(* CODESYS project keyence_iv.library
   Company: KOSTAL GmbH & Co.KG
   Version: 2.0.0.0
   DefaultNamespace: KOSTAL.AF2024.Drivers.Camera.Keyence_IV
   Title: KOSTAL.AF2024.Drivers.Camera.Keyence_IV
   Placeholder: KOSTAL.AF2024.Drivers.Camera.Keyence_IV
   Author: Frank Dümpelmann, Martin Hundt
   DocFormat: reStructuredText

Project tree, tasks and I/O mapping:
  libraries: KOSTAL.AF2024.Core.functionResponse, 1.0.0.0 (KOSTAL GmbH & Co.KG); KOSTAL.AF2024.Core.ListOf, 1.0.0.0 (KOSTAL GmbH & Co.KG); KOSTAL.AF2024.Core.Process, 1.0.0.0 (KOSTAL GmbH & Co.KG); KOSTAL.AF2024.Core.Settings, 1.0.0.0 (KOSTAL GmbH & Co.KG); KOSTAL.AF2024.Core.StringTools, 1.0.0.0 (KOSTAL GmbH & Co.KG); KOSTAL.AF2024.Core.System, 1.0.0.0 (KOSTAL GmbH & Co.KG); KOSTAL.AF2024.Drivers.Camera.I_Camera, 2.0.0.0 (KOSTAL GmbH & Co.KG); Tc2_Standard, 3.3.3.0 (Beckhoff Automation GmbH); Tc2_System, 3.6.2.0 (Beckhoff Automation GmbH); Tc2_TcpIp, 3.3.10.0 (Beckhoff Automation GmbH)
  DIO/
    DUT/
      data type _E_PROCESS
      data type _ST_fromDevice
      data type _ST_fromDevice_HG_
      data type _ST_toDevice
    function block FB_Camera_DIO_IV [ST]: Ex_SetProgramNumber, Ex_Trigger, Ex_Trigger_ProgramNumber, ProgramNumber, ResultPass, State, _setFinish, _toDevice_Clear, _faultHandler, _fbMain, _idle, _sequence, _setProgram, Fault, FaultReset, FBmain
    function block FB_Camera_DIO_IV_HG [ST]: CustomOut_5, CustomOut_6, CustomOut_7, CustomOut_8
  Project Information/
    function F_GetCompany [ST]
    function F_GetTitle [ST]
    function F_GetVersion [ST]
  TcpIp/
    DUT/
      _Internal/
        data type _E_Command_TcpIp
        data type _E_THIS_TcpIp
        function block _T_Command [ST]: Error, GetProgram, OK, ReadOperationMode, ReadVersion, SetProgram, StateResult, TriggerAndState
      Response RT/
        interface I_T_Response_RT_TcpIp: CopyTo, OverallPass, ResultCount, Tools
        interface I_T_Response_RT_TcpIp_CopyFrom: CopyFrom
        interface I_T_Response_RT_TcpIp_Owner: Clear, CopyFrom, OverallPass, ResultCount, Tools_Owner
        function block T_Response_RT_TcpIp [ST]: Clear, CopyFrom, CopyTo, OverallPass, ResultCount, Tools, Tools_Owner
      Tool/
        ListOf/
          function block FB_ListOf_T_Tool [ST]: _get_I, _get_I_Owner, _removePayLoad, _verifyMember, Add_DUT, Clear, CopyFrom, CopyTo, Delete_DUT, Get_I, Get_I_Owner, NumberOfMember
          interface I_ListOf_T_Tool: CopyTo, Get_I, NumberOfMember
          interface I_ListOf_T_Tool_CopyFrom: CopyFrom
          interface I_ListOf_T_Tool_Owner: Add_DUT, Clear, CopyFrom, CopyTo, Delete_DUT, Get_I, Get_I_Owner, NumberOfMember
        interface I_T_Tool: CopyTo, MatchingRate, Number, Pass
        interface I_T_Tool_CopyFrom: CopyFrom
        interface I_T_Tool_Owner: Clear, CopyFrom, MatchingRate, Number, Pass
        function block T_Tool [ST]: Clear, CopyFrom, CopyTo, MatchingRate, Number, Pass
      Version/
        interface I_T_SensorVersion_TcpIp: CopyTo, HeadModel, Version
        interface I_T_SensorVersion_TcpIp_CopyFrom: CopyFrom
        interface I_T_SensorVersion_TcpIp_Owner: Clear, CopyFrom, HeadModel, Version
        function block T_SensorVersion_TcpIp [ST]: Clear, CopyFrom, CopyTo, HeadModel, Version
      data type E_OpMode_TcpIp
    function block FB_Camera_TcpIp_IV [ST]: FB_init, _getCommand, _mergePlCommand, _Parse_Error, _Parse_ErrorMessage, _Parse_GetProgram, _Parse_OpMode, _Parse_SetProgram, _Parse_Trigger, _Parse_Version, _a0_stepFail, _a0_stepInit, _a1_Finish, _a1_Idle, _a2_Connect, _a2_Parse, _a2_Receive, _a2_Send, _a3_PrgIsEqual, _devices, _splitString, _timeOutOccured, _FBmain, Clear, Ex_GetProgramNumber, Ex_ReadOperationMode, Ex_ReadVersion, Ex_SetProgramNumber, Ex_Trigger, Ex_Trigger_ProgramNumber, GetElement, NativeStringGet, IP, Port, Content, ExecutedSocketState, NumberOfEntries, OperationMode, Result, ResultPass, serverAmsNetId, State, Version, FBmain
    interface I_Camera_TcpIp_IV: GetElement, NativeStringGet, Content, ExecutedSocketState, IP, NumberOfEntries, OperationMode, Port, Result, serverAmsNetId
  Version/
    global variables Global_Version
*)

// DIO/DUT/_E_PROCESS
{attribute 'qualified_only'}
{attribute 'strict'}
TYPE _E_PROCESS :
(
	idle		:= 0,
	Start		:= 1, 
	SetProgram	:= 2
);
END_TYPE

// DIO/DUT/_ST_fromDevice
TYPE _ST_fromDevice :
STRUCT
	TotalStatusOK	:BOOL;
	Busy			:BOOL;
	Error			:BOOL;
	Run				:BOOL;
END_STRUCT
END_TYPE

// DIO/DUT/_ST_fromDevice_HG_
TYPE _ST_fromDevice_HG_ :
STRUCT
	CustomOut_5		: BOOL;
	CustomOut_6		: BOOL;
	CustomOut_7		: BOOL;
	CustomOut_8		: BOOL;
END_STRUCT
END_TYPE

// DIO/DUT/_ST_toDevice
TYPE _ST_toDevice:
	STRUCT
		ExternalTrigger		:BOOL;
		ProgramSelectBit0	:BOOL;
		ProgramSelectBit1	:BOOL;
		ProgramSelectBit2	:BOOL;
		ProgramSelectBit3	:BOOL;
		ErrorClear			:BOOL;
	END_STRUCT
END_TYPE

// TcpIp/DUT/_Internal/_E_Command_TcpIp
{attribute 'qualified_only'}
{attribute 'strict'}
TYPE INTERNAL _E_Command_TcpIp :
(
	Trigger := 0,
	SetProgram,
	GetProgram,
	ReadVersion,
	ReadOperationMode
);
END_TYPE

// TcpIp/DUT/_Internal/_E_THIS_TcpIp
{attribute 'qualified_only'}
{attribute 'strict'}
TYPE INTERNAL _E_THIS_TcpIp :
(
	Idle := 0,
	Trigger,
	TriggerPrgNo,
	SetProgram,
	GetProgram,
	ReadVersion,
	ReadOperationMode
);
END_TYPE

// TcpIp/DUT/E_OpMode_TcpIp
{attribute 'qualified_only'}
{attribute 'strict'}
TYPE E_OpMode_TcpIp :
(
	Unknown := 0,
	Setup,
	Run
);
END_TYPE

// Version/Global_Version
{attribute 'TcGenerated'}
{attribute 'no-analysis'}
{attribute 'linkalways'}
// This function has been automatically generated from the project information.
VAR_GLOBAL CONSTANT
	{attribute 'const_non_replaced'}
	stLibVersion_KOSTAL_AF2024_Drivers_Camera_Keyence_IV : ST_LibVersion := (iMajor := 2, iMinor := 0, iBuild := 0, iRevision := 0, nFlags := 0, sVersion := '2.0.0.0');
END_VAR

// DIO/FB_Camera_DIO_IV
(*

:Author: Martin Hundt <m.hundt@kostal.com>
:Date: 2022-03-11

Function
========
| Device driver for Keyence IV-Series vision sensors with discrete IOs
| Selection of 15 sensor programs (program No. 0 is reserved)

Methods and Properties
======================
| Ex_start: Start the last selected camera program
| Ex_start_ProgramNumber: Start the camera program number in the method's parameter (int)

| State.ready: Camera is ready
| State.busy: Camera is analysing an image
| State.finish: Image analysis was finished
| State.pass: Image was processed -> Check result
| State.fail: Image image processing failed

| Fault: Camera in error state


Sensor Configuration
=====================
| The following IOs must be configured at the sensor and linked to the hardware IOs according to their names:
| Sensor Outputs: TotalStatusOK, Busy, Error, Run				
| Sensor Inputs: ExternalTrigger, ProgramSelectBit0, ProgramSelectBit1, ProgramSelectBit2, ErrorClear			

*)

FUNCTION_BLOCK FB_Camera_DIO_IV IMPLEMENTS KOSTAL_AF2024_Drivers_Camera_I_Camera.I_CameraWithFeedback
VAR
	_fromSensor AT %I*	: _ST_fromDevice;
	_toSensor 	AT %Q*	: _ST_toDevice;
	
	_THIS_CALLED		: _E_PROCESS;
	_THIS_IN_PROCESS	: _E_PROCESS;
	_step				: KOSTAL_AF2024_Core_Process.FB_processStep;
	_state				: KOSTAL_AF2024_Core_Process.T_plcState;
	
	_programNoOld		: USINT;
	_init				: BOOL;		(*BOOL - initialization required*)
	_triggerBusy		: F_TRIG;	(*F_TRIG*)
	_responseTime		: TON;	(*TON*)
	_resetClock			: TP;		(*TP*)
	
	_faultReset			: BOOL;
	
	_resultPass			: BOOL;
	_resultFail			: BOOL;
	
	_programNo			: USINT;
	_fault				: BOOL;
	                    
END_VAR

METHOD Ex_SetProgramNumber : BOOL;
VAR_INPUT
	ProgramNumber	: UINT;
END_VAR
IF _THIS_CALLED <> _E_PROCESS.idle THEN //Another process is running: don't start this process!
	Ex_SetProgramNumber:= FALSE;	
	RETURN; 
END_IF

_programNo := UINT_TO_USINT(ProgramNumber);
_THIS_CALLED := _E_PROCESS.SetProgram;

_FBmain();	//Call sequence via _FBmain

Ex_SetProgramNumber := _THIS_CALLED = _THIS_IN_PROCESS;	//Return true when process was started
END_METHOD

METHOD Ex_Trigger : BOOL;
IF _THIS_CALLED <> _E_PROCESS.idle THEN //Another process is running: don't start this process!
	Ex_Trigger:= FALSE;	
	RETURN; 
END_IF


_THIS_CALLED := _E_PROCESS.Start;

_FBmain();	//Call sequence via _FBmain

Ex_Trigger := _THIS_CALLED = _THIS_IN_PROCESS;	//Return true when process was started
END_METHOD

METHOD Ex_Trigger_ProgramNumber : BOOL;
VAR_INPUT
	ProgramNumber	: UINT;
END_VAR
IF _THIS_CALLED <> _E_PROCESS.idle THEN //Another process is running: don't start this process!
	Ex_Trigger_ProgramNumber:= FALSE;	
	RETURN; 
END_IF

_programNo := UINT_TO_USINT(ProgramNumber);
_THIS_CALLED := _E_PROCESS.Start;

_FBmain();	//Call sequence via _FBmain

Ex_Trigger_ProgramNumber := _THIS_CALLED = _THIS_IN_PROCESS;	//Return true when process was started
END_METHOD

PROPERTY PUBLIC ProgramNumber : UINT
GET
ProgramNumber := _programNo;
END_GET
END_PROPERTY

PROPERTY PUBLIC ResultPass : BOOL
GET
ResultPass := _resultPass;
END_GET
END_PROPERTY

PROPERTY State : KOSTAL_AF2024_Core_Process.I_T_plcState
GET

State := _state;
END_GET
END_PROPERTY

METHOD PROTECTED _setFinish
VAR_INPUT
END_VAR
END_METHOD

METHOD PROTECTED _toDevice_Clear
VAR_INPUT
END_VAR
_toSensor.ErrorClear := FALSE;
_toSensor.ExternalTrigger := FALSE;
_toSensor.ProgramSelectBit0 := FALSE;
_toSensor.ProgramSelectBit1 := FALSE;
_toSensor.ProgramSelectBit2 := FALSE;
_toSensor.ProgramSelectBit3 := FALSE;
END_METHOD

METHOD PROTECTED _faultHandler : BOOL
VAR_INPUT
END_VAR
_fault:= _fromSensor.Error;

IF _fromSensor.Error THEN
	_state.clear();
	_state.Fail:= TRUE;
	_state.Description:= "Device send >ERROR<";	
	
	_toDevice_Clear();

	_resetClock(IN:= _faultReset, PT:= T#250MS);
	_toSensor.ErrorClear:= _resetClock.Q;	
ELSE
	_faultHandler := TRUE;
END_IF

_faultReset := false;
END_METHOD

METHOD Protected _fbMain
VAR_INPUT
END_VAR
IF NOT _init THEN
	_step.init();
	_programNoOld:= 0;
	_resetClock(IN:= FALSE);
	_init:= TRUE;
	_toDevice_Clear();
END_IF

IF NOT _faultHandler() THEN RETURN; END_IF


IF _THIS_CALLED <> _THIS_IN_PROCESS THEN
	_step.init();
END_IF

_THIS_IN_PROCESS:= _THIS_CALLED;

CASE _THIS_CALLED OF
	_E_PROCESS.SetProgram:
		_setProgram();
	_E_PROCESS.Start:
		_sequence();
ELSE
	_idle();
END_CASE
END_METHOD

METHOD PROTECTED _idle
VAR_INPUT
END_VAR
_step.init();

_toSensor.ErrorClear:= FALSE;
_toSensor.ExternalTrigger := FALSE;
_resultPass := FALSE;
_resultFail := FALSE;
_state.clear();
_state.Ready := TRUE;
END_METHOD

METHOD PROTECTED _sequence
VAR_INPUT
END_VAR
_step.Header();

CASE _step.actual OF		
	0: //Check Program No.
		_state.clear();
		_state.Busy := TRUE;
		IF (_programNo = 0) OR (_programNo > 15) THEN
			_state.clear();
			_state.finish:= TRUE;
			_state.Fail:= TRUE;
			_state.Description:= "ProgramNo out of range (1<Pno>15)";
		ELSE
			_step.INC();
		END_IF

	1: (*Change Program *)
		IF _step.Toggle THEN
			_responseTime(IN:= FALSE);
			_triggerBusy(CLK:= FALSE);
		END_IF

		_toSensor.ProgramSelectBit0 := _programNo.0;
		_toSensor.ProgramSelectBit1 := _programNo.1;
		_toSensor.ProgramSelectBit2 := _programNo.2;
		_toSensor.ProgramSelectBit3 := _programNo.3;

		_state.clear();
		_state.Busy := TRUE;
		_state.Description:= "send program Number";

		_responseTime(IN:= TRUE, PT:= T#1s);
		_triggerBusy(CLK:=_fromSensor.Busy);	(*Wait until program is changed*)

		IF _programNo <> _programNoOld THEN

			IF _triggerBusy.Q OR _responseTime.Q THEN
				_programNoOld := _programNo;
			END_IF

		ELSE
			_step.INC();
		END_IF

	2:	(*trigger*)
		_toSensor.ExternalTrigger := TRUE;

		_state.clear();
		_state.Busy := TRUE;
		_state.Description:= "wait sensor busy";

		IF NOT _fromSensor.Run THEN
			_state.clear();
			_state.finish := TRUE;
			_state.fail := TRUE;
			_state.Description:= "Device not in >RUN<";
		ELSIF _fromSensor.Busy THEN
			_step.INC();
		END_IF

	3:	(*Read result*)
		_toSensor.ExternalTrigger := TRUE;

		_state.clear();
		_state.Busy := TRUE;
		_state.Description:=  "wait sensor finish";

		IF NOT _fromSensor.Busy THEN
			_step.INC();
		END_IF

	4:	(*finish*)
		_toSensor.ExternalTrigger := TRUE;
		_state.clear();
		_state.Finish := TRUE;
		_state.pass := TRUE;
		
		_resultPass:= _fromSensor.TotalStatusOK;
		_resultFail:= NOT _fromSensor.TotalStatusOK;

		
		IF _resultPass THEN
			_state.Description:= "get PASS";
		ELSE
			_state.Description:= "get FAIL";
		END_IF
		

END_CASE
END_METHOD

METHOD PROTECTED _setProgram
VAR_INPUT
END_VAR
_state.clear();
IF (_programNo = 0) OR (_programNo > 15) THEN
	_state.finish:= TRUE;
	_state.Fail:= TRUE;
	_state.Description:= "ProgramNo out of range (1<Pno>15)";
ELSE
	_state.finish:= TRUE;
	_state.pass:= TRUE;
END_IF
END_METHOD

PROPERTY Fault : BOOL
GET
Fault := _fault;
END_GET
END_PROPERTY

METHOD PUBLIC FaultReset
VAR_INPUT
END_VAR
_faultReset := True;
END_METHOD

METHOD PUBLIC FBmain
VAR_INPUT
END_VAR
IF _THIS_CALLED = _E_PROCESS.idle THEN
	
	_FBmain();
	
END_IF

_THIS_CALLED:= _E_PROCESS.idle;
END_METHOD

END_FUNCTION_BLOCK

// DIO/FB_Camera_DIO_IV_HG
//Extension of FB_Camera_IV with four custom outputs (only available for IV-HG device)
FUNCTION_BLOCK FB_Camera_DIO_IV_HG EXTENDS FB_Camera_DIO_IV
VAR
	_fromdeviceCustom	AT %I*	: _ST_fromDevice_HG_;
END_VAR

PROPERTY PUBLIC CustomOut_5 : Bool
GET
CustomOut_5 := _fromdeviceCustom.CustomOut_5;
END_GET
END_PROPERTY

PROPERTY PUBLIC CustomOut_6 : Bool
GET
CustomOut_6 := _fromdeviceCustom.CustomOut_6;
END_GET
END_PROPERTY

PROPERTY PUBLIC CustomOut_7 : Bool
GET
CustomOut_7 := _fromdeviceCustom.CustomOut_7;
END_GET
END_PROPERTY

PROPERTY PUBLIC CustomOut_8 : Bool
GET
CustomOut_8 := _fromdeviceCustom.CustomOut_8;
END_GET
END_PROPERTY

END_FUNCTION_BLOCK

// Project Information/F_GetCompany
// This function has been automatically generated from the project information.
{attribute 'signature_flag' := '1073741824'}
{attribute 'TcGenerated'}
{attribute 'no-analysis'}
FUNCTION F_GetCompany : WSTRING
VAR_INPUT
	
END_VAR

F_GetCompany := "KOSTAL GmbH & Co.KG";

END_FUNCTION

// Project Information/F_GetTitle
// This function has been automatically generated from the project information.
{attribute 'signature_flag' := '1073741824'}
{attribute 'TcGenerated'}
{attribute 'no-analysis'}
FUNCTION F_GetTitle : WSTRING
VAR_INPUT
	
END_VAR

F_GetTitle := "KOSTAL.AF2024.Drivers.Camera.Keyence_IV";

END_FUNCTION

// Project Information/F_GetVersion
// This function has been automatically generated from the project information.
{attribute 'signature_flag' := '1073741824'}
{attribute 'TcGenerated'}
{attribute 'no-analysis'}
FUNCTION F_GetVersion : ST_LibVersion
VAR_INPUT
	
END_VAR

F_GetVersion.iMajor := 2;
F_GetVersion.iMinor := 0;
F_GetVersion.iBuild := 0;
F_GetVersion.iRevision := 0;
F_GetVersion.sVersion := '2.0.0.0';
F_GetVersion.nFlags := 0;

END_FUNCTION

// TcpIp/DUT/_Internal/_T_Command
FUNCTION_BLOCK INTERNAL _T_Command

PROPERTY PUBLIC Error : STRING
GET

Error	:= 'ER';
END_GET
END_PROPERTY

PROPERTY PUBLIC GetProgram : STRING
GET

GetProgram	:= 'PR';
END_GET
END_PROPERTY

PROPERTY PUBLIC OK : STRING
GET

OK	:= 'OK';
END_GET
END_PROPERTY

PROPERTY PUBLIC ReadOperationMode : STRING
GET

ReadOperationMode	:= 'RM';
END_GET
END_PROPERTY

PROPERTY PUBLIC ReadVersion : STRING
GET

ReadVersion	:= 'VI';
END_GET
END_PROPERTY

PROPERTY PUBLIC SetProgram : STRING
GET

SetProgram	:= 'PW';
END_GET
END_PROPERTY

PROPERTY PUBLIC StateResult : STRING
GET

StateResult	:= 'RT';
END_GET
END_PROPERTY

PROPERTY PUBLIC TriggerAndState : STRING
GET

TriggerAndState	:= 'T2';
END_GET
END_PROPERTY

END_FUNCTION_BLOCK

// TcpIp/DUT/Response RT/I_T_Response_RT_TcpIp
INTERFACE I_T_Response_RT_TcpIp EXTENDS KOSTAL_AF2024_Core_System.I_Interface

METHOD PUBLIC CopyTo : BOOL
VAR_INPUT
	IN	: I_T_Response_RT_TcpIp_CopyFrom;
END_VAR
END_METHOD

PROPERTY PUBLIC OverallPass : BOOL
GET
END_GET
END_PROPERTY

PROPERTY PUBLIC ResultCount : UDINT
GET
END_GET
END_PROPERTY

PROPERTY PUBLIC Tools : I_ListOf_T_Tool
GET
END_GET
END_PROPERTY

END_INTERFACE

// TcpIp/DUT/Response RT/I_T_Response_RT_TcpIp_CopyFrom
INTERFACE I_T_Response_RT_TcpIp_CopyFrom EXTENDS KOSTAL_AF2024_Core_System.I_Interface

METHOD PUBLIC CopyFrom : BOOL
VAR_INPUT
	IN	: I_T_Response_RT_TcpIp;
END_VAR
END_METHOD

END_INTERFACE

// TcpIp/DUT/Tool/ListOf/I_ListOf_T_Tool
(*
	Read only Interface from List of DUT
*)
INTERFACE I_ListOf_T_Tool EXTENDS KOSTAL_AF2024_Core_ListOf._I_Object_Base

METHOD PUBLIC CopyTo : BOOL
VAR_INPUT
	IN	: I_ListOf_T_Tool_CopyFrom;
END_VAR
END_METHOD

METHOD Get_I : BOOL

VAR_INPUT
	Number		: UDINT;
	rFound_I	: REFERENCE TO I_T_Tool;
	Response	: KOSTAL_AF2024_Core_functionResponse.I_T_functionResponse_Owner;
END_VAR
END_METHOD

PROPERTY NumberOfMember : UDINT
GET
END_GET
END_PROPERTY

END_INTERFACE

// TcpIp/DUT/Tool/ListOf/I_ListOf_T_Tool_CopyFrom
(*
	The class implementing this interface can take over the contents from another instance with the same interface {I_DUT}.
	Typing takes place in the method.
*)
INTERFACE I_ListOf_T_Tool_CopyFrom EXTENDS KOSTAL_AF2024_Core_System.I_Interface

(*
	Copies the contents of another list {IN} into its own memory.
*)
METHOD PUBLIC CopyFrom : BOOL
VAR_INPUT
	IN	: KOSTAL_AF2024_Core_System.I_Interface;
END_VAR
END_METHOD

END_INTERFACE

// TcpIp/DUT/Tool/I_T_Tool
(*
	Read only Interface from DUT
*)
INTERFACE I_T_Tool  EXTENDS KOSTAL_AF2024_Core_System.I_Interface

METHOD PUBLIC CopyTo : bool
VAR_INPUT
	IN	: I_T_Tool_CopyFrom;
END_VAR
END_METHOD

PROPERTY PUBLIC MatchingRate : KOSTAL_AF2024_Core_Settings.T_MaxString_UTF8
GET
END_GET
END_PROPERTY

PROPERTY PUBLIC Number : UINT
GET
END_GET
END_PROPERTY

PROPERTY PUBLIC Pass : BOOL
GET
END_GET
END_PROPERTY

END_INTERFACE

// TcpIp/DUT/Tool/I_T_Tool_CopyFrom
INTERFACE I_T_Tool_CopyFrom EXTENDS KOSTAL_AF2024_Core_System.I_Interface

METHOD PUBLIC CopyFrom : BOOL
VAR_INPUT
	IN	: KOSTAL_AF2024_Core_System.I_Interface;
END_VAR
END_METHOD

END_INTERFACE

// TcpIp/DUT/Response RT/I_T_Response_RT_TcpIp_Owner
INTERFACE I_T_Response_RT_TcpIp_Owner EXTENDS I_T_Response_RT_TcpIp

METHOD PUBLIC Clear
VAR_INPUT
END_VAR
END_METHOD

METHOD PUBLIC CopyFrom : BOOL
VAR_INPUT
	IN	: I_T_Response_RT_TcpIp;
END_VAR
END_METHOD

PROPERTY PUBLIC OverallPass : BOOL
SET
END_SET
END_PROPERTY

PROPERTY PUBLIC ResultCount : UDINT
SET
END_SET
END_PROPERTY

PROPERTY PUBLIC Tools_Owner : I_ListOf_T_Tool_Owner
GET
END_GET
END_PROPERTY

END_INTERFACE

// TcpIp/DUT/Tool/ListOf/I_ListOf_T_Tool_Owner
(*
	Full qualified access Interface from List of DUT
*)
INTERFACE I_ListOf_T_Tool_Owner EXTENDS KOSTAL_AF2024_Core_ListOf._I_Object_Base_Owner

//Add a new instance of FB_Dut and copy content from [IN] to the new instance
METHOD PUBLIC Add_DUT : BOOL
VAR_INPUT
	IN				: KOSTAL_AF2024_Core_System.I_Interface;
	Response	: KOSTAL_AF2024_Core_functionResponse.I_T_functionResponse_Owner;
END_VAR
END_METHOD

METHOD Clear
VAR_INPUT
END_VAR
END_METHOD

METHOD PUBLIC CopyFrom : BOOL
VAR_INPUT
	IN	: KOSTAL_AF2024_Core_System.I_Interface;
END_VAR
END_METHOD

METHOD PUBLIC CopyTo : BOOL
VAR_INPUT
	IN	: I_ListOf_T_Tool_CopyFrom;
END_VAR
END_METHOD

METHOD PUBLIC Delete_DUT : BOOL
VAR_INPUT
	Number	: UDINT;	//Number of DUT in List
	Response	: KOSTAL_AF2024_Core_functionResponse.I_T_functionResponse_Owner;
END_VAR
END_METHOD

METHOD Get_I : BOOL

VAR_INPUT
	Number		: UDINT;
	rFound_I	: REFERENCE TO I_T_Tool;
	Response	: KOSTAL_AF2024_Core_functionResponse.I_T_functionResponse_Owner;
END_VAR
END_METHOD

//Get full access to content 
METHOD Get_I_Owner : BOOL

VAR_INPUT
	Number		: UDINT;
	rFound_I	: REFERENCE TO I_T_Tool_Owner;
	Response	: KOSTAL_AF2024_Core_functionResponse.I_T_functionResponse_Owner;
END_VAR
END_METHOD

PROPERTY NumberOfMember : UDINT
GET
END_GET
END_PROPERTY

END_INTERFACE

// TcpIp/DUT/Tool/I_T_Tool_Owner
(*
	Full qualified access Interface from DUT
*)
INTERFACE I_T_Tool_Owner EXTENDS I_T_Tool

METHOD PUBLIC Clear
VAR_INPUT
END_VAR
END_METHOD

METHOD PUBLIC CopyFrom : BOOL
VAR_INPUT
	IN	: KOSTAL_AF2024_Core_System.I_Interface;
END_VAR
END_METHOD

PROPERTY PUBLIC MatchingRate : KOSTAL_AF2024_Core_Settings.T_MaxString_UTF8
SET
END_SET
END_PROPERTY

PROPERTY PUBLIC Number : UINT
SET
END_SET
END_PROPERTY

PROPERTY PUBLIC Pass : BOOL
SET
END_SET
END_PROPERTY

END_INTERFACE

// TcpIp/DUT/Response RT/T_Response_RT_TcpIp
FUNCTION_BLOCK PUBLIC T_Response_RT_TcpIp IMPLEMENTS I_T_Response_RT_TcpIp, I_T_Response_RT_TcpIp_Owner, I_T_Response_RT_TcpIp_CopyFrom

VAR
	_ResultCount	: UDINT;
	_OverallPass	: BOOL;
	_Tools				: FB_ListOf_T_Tool;
END_VAR

METHOD PUBLIC Clear
VAR_INPUT
END_VAR

_ResultCount	:= UDINT#0;
_OverallPass	:= FALSE;
_Tools.Clear();
END_METHOD

METHOD PUBLIC CopyFrom : BOOL
VAR_INPUT
	IN	: I_T_Response_RT_TcpIp;
END_VAR

VAR
	_obj	: I_T_Response_RT_TcpIp;
END_VAR

IF (IN = 0) OR_ELSE NOT __QUERYINTERFACE(IN, _obj) OR_ELSE (_obj = 0) THEN RETURN;	END_IF

_OverallPass	:= IN.OverallPass;
_ResultCount	:= IN.ResultCount;
_Tools.CopyFrom(IN.Tools);

CopyFrom:= TRUE;
END_METHOD

METHOD PUBLIC CopyTo : BOOL
VAR_INPUT
	IN	: I_T_Response_RT_TcpIp_CopyFrom;
END_VAR

VAR
	_obj	: I_T_Response_RT_TcpIp_CopyFrom;
END_VAR

IF (IN = 0) OR_ELSE NOT __QUERYINTERFACE(IN, _obj) OR_ELSE (_obj = 0) THEN RETURN;	END_IF

CopyTo:= IN.CopyFrom(THIS^);
END_METHOD

PROPERTY PUBLIC OverallPass : BOOL
GET

OverallPass:= _OverallPass;
END_GET
SET

_OverallPass:= OverallPass;
END_SET
END_PROPERTY

PROPERTY PUBLIC ResultCount : UDINT
GET

ResultCount:= _ResultCount;
END_GET
SET

_ResultCount:= ResultCount;
END_SET
END_PROPERTY

PROPERTY PUBLIC Tools : I_ListOf_T_Tool
GET

Tools:= _Tools;
END_GET
END_PROPERTY

PROPERTY PUBLIC Tools_Owner : I_ListOf_T_Tool_Owner
GET

Tools_Owner:= _Tools;
END_GET
END_PROPERTY

END_FUNCTION_BLOCK

// TcpIp/DUT/Tool/ListOf/FB_ListOf_T_Tool
(*
	A template for creating a list of typed classes (FBs)
*)
FUNCTION_BLOCK FB_ListOf_T_Tool EXTENDS KOSTAL_AF2024_Core_ListOf._FB_Object_Base  IMPLEMENTS I_ListOf_T_Tool, I_ListOf_T_Tool_CopyFrom, I_ListOf_T_Tool_Owner

VAR
	//Use the {_Dummy} to ensure that a valid interface is always returned.
	_Dummy	: T_Tool;
END_VAR

(*
	Returns the typed interface in the reference variable.
	In the event of an error, the return value becomes FALSE and the interface refers to the {_Dummy}.
*)
METHOD PROTECTED _get_I : BOOL

VAR_INPUT
	Member		: KOSTAL_AF2024_Core_System.I_Interface;
	rFound_I	: REFERENCE TO I_T_Tool;
	Response	: KOSTAL_AF2024_Core_functionResponse.I_T_functionResponse_Owner;
END_VAR

VAR
	_iObj			: I_T_Tool;
	_Success	: BOOL;
END_VAR
//preset
IF 		__ISVALIDREF(rFound_I)	THEN	rFound_I:= _Dummy;	
ELSE 	_setResultFail(Response, "no reference to rFound_I found");	RETURN; 
END_IF	

IF NOT _verifyMember(Member, Response)	THEN RETURN;	END_IF

_Success:= __QUERYINTERFACE(Member, _iObj);

//return dummy if no valid DUT is found
IF NOT _Success OR_ELSE (_iObj = 0)	THEN	
	_setResultFail(Response, "__QueryInterface failed - return Dummy");	RETURN;	
END_IF

rFound_I:= _iObj;
_setResultPass(Response, "Successful");

_get_I:= TRUE;
END_METHOD

(*
	Returns the typed owner interface in the reference variable.
	In the event of an error, the return value becomes FALSE and the interface refers to the {_Dummy}.
*)
METHOD PROTECTED _get_I_Owner : BOOL

VAR_INPUT
	Member		: KOSTAL_AF2024_Core_System.I_Interface;
	rFound_I	: REFERENCE TO I_T_Tool_Owner;
	Response	: KOSTAL_AF2024_Core_functionResponse.I_T_functionResponse_Owner;
END_VAR

VAR
	_iObj			: I_T_Tool_Owner;
	_Success	: BOOL;
END_VAR
//preset
IF 		__ISVALIDREF(rFound_I)	THEN	rFound_I:= _Dummy;	
ELSE 	_setResultFail(Response, "no reference to rFound_I found");	RETURN; 
END_IF	

IF NOT _verifyMember(Member, Response)	THEN RETURN;	END_IF

_Success:= __QUERYINTERFACE(Member, _iObj);

//return dummy if no valid DUT is found
IF NOT _Success OR_ELSE (_iObj = 0)	THEN	
	_setResultFail(Response, "__QueryInterface failed - return Dummy");	RETURN;	
END_IF

rFound_I:= _iObj;
_setResultPass(Response, "Successful");

_get_I_Owner:= TRUE;
END_METHOD

(*
	Cleans the custom class {FB_DUT} and removes it from memory.
*)
METHOD PROTECTED  _removePayLoad : BOOL
VAR_INPUT
	Member	: KOSTAL_AF2024_Core_System.I_Interface;
	Result	: KOSTAL_AF2024_Core_functionResponse.I_T_functionResponse_Owner;
END_VAR

VAR
	_iObj			: I_T_Tool_Owner;
	_pFB_DUT	:	POINTER TO T_Tool;
	_Success	: BOOL;
END_VAR


IF NOT SUPER^._removePayload(Member, Result)	THEN RETURN;	END_IF

_Success:= __QUERYINTERFACE(Member, _iObj);

IF NOT _Success	THEN	RETURN;	END_IF
IF _iObj = 0		THEN	RETURN;	END_IF

_iObj.Clear();

_Success  := __QUERYPOINTER(_iObj, _pFB_DUT);

IF NOT _Success	THEN	RETURN;	END_IF
IF _pFB_DUT = 0	THEN	RETURN;	END_IF

__DELETE(_pFB_DUT);
END_METHOD

(*
	Overload the method from the base class to verify the custom interface. 
	The local method {_get_I_Owner()} is used for this.
*)
METHOD PROTECTED _verifyMember : BOOL

VAR_INPUT
	Member	: KOSTAL_AF2024_Core_System.I_Interface;
	Result	: KOSTAL_AF2024_Core_functionResponse.I_T_functionResponse_Owner;
END_VAR

VAR
	_pObj	: POINTER TO T_Tool;
	_Success: BOOL;
END_VAR

IF NOT SUPER^._verifyMember(Member, Result)	THEN RETURN;	END_IF

_Success:= __QUERYPOINTER(Member, _pObj);

//return dummy if no valid Pointer to DUT is found
IF NOT _Success OR_ELSE (_pObj = 0)	THEN	_setResultFail(Result, "__QueryInterface failed");	RETURN; END_IF

_verifyMember:= TRUE;
END_METHOD

(*
	Add a new instance of FB_Dut and copy content from [IN] to the new instance
*)
METHOD PUBLIC Add_DUT : BOOL
VAR_INPUT
	IN				: KOSTAL_AF2024_Core_System.I_Interface;
	Response	: KOSTAL_AF2024_Core_functionResponse.I_T_functionResponse_Owner;
END_VAR

VAR
	_pDUT: POINTER TO T_Tool;
END_VAR

_pDUT:= __NEW(T_Tool);

IF _pDUT = 0 THEN	_setResultFail(Response, "cannot create new object"); RETURN; END_IF

IF NOT _pDUT^.CopyFrom(IN) THEN
	
	_setResultFail(Response, "cannot copy content");

	__DELETE(_pDUT);

	RETURN;

END_IF

Add_DUT:= _addMember(_pDUT^, Response);
END_METHOD

(*
	Makes the protected method public.
*)
METHOD Clear

_clear();
END_METHOD

(*
	Copies the contents of another list {IN} into its own memory.
*)
METHOD PUBLIC CopyFrom : BOOL
VAR_INPUT
	IN	: KOSTAL_AF2024_Core_System.I_Interface;
END_VAR

VAR
	_udi	: UDINT;

	_obj	: I_ListOf_T_Tool;
	_IDUT	: I_T_Tool;

	_obj2		: I_ListOf_T_Tool_Owner;
	_IDUT2	: I_T_Tool_Owner;
END_VAR
_clear();

IF IN = 0 THEN RETURN;

ELSIF __QUERYINTERFACE(IN, _obj) AND_THEN _obj <> 0 THEN
	
	FOR _udi:= 1 TO _obj.NumberOfMember DO
		IF _obj.Get_I(_udi, _IDUT, 0)	THEN	Add_DUT(_IDUT, 0);	END_IF
	END_FOR

	CopyFrom:= TRUE;

ELSIF __QUERYINTERFACE(IN, _obj2) AND_THEN _obj2 <> 0 THEN
	
	FOR _udi:= 1 TO _obj2.NumberOfMember DO
		IF _obj2.Get_I_Owner(_udi, _IDUT2, 0)	THEN	Add_DUT(_IDUT2, 0);	END_IF
	END_FOR

	CopyFrom:= TRUE;

END_IF
END_METHOD

(*
	Copies the own content into another list created at the parameter {IN}.
*)
METHOD PUBLIC CopyTo : BOOL
VAR_INPUT
	IN	: I_ListOf_T_Tool_CopyFrom;
END_VAR

IF IN = 0 THEN RETURN;	END_IF

CopyTo:= IN.CopyFrom(THIS^);
END_METHOD

(*
	Deletes the class specified with the {Number} from the list.
*)
METHOD PUBLIC Delete_DUT : BOOL
VAR_INPUT
	Number		: UDINT;	//Number of DUT in List
	Response	: KOSTAL_AF2024_Core_functionResponse.I_T_functionResponse_Owner;
END_VAR

VAR
	//_response	: KOSTAL_AF2024_Core_functionResponse.T_functionResponse;
	_Success	: BOOL;
	_Member		: KOSTAL_AF2024_Core_System.I_Interface;
END_VAR

IF Number = 0 THEN	_setResultFail(Response, "Number is out of range (1..n)"); RETURN; END_IF

Delete_DUT:= _removeMemberByIndex(Number - 1, Response);
END_METHOD

(*
	Get readonly access to content of Member with {Number}
*) 
METHOD Get_I : BOOL

VAR_INPUT
	Number		: UDINT;
	rFound_I	: REFERENCE TO I_T_Tool;
	Response	: KOSTAL_AF2024_Core_functionResponse.I_T_functionResponse_Owner;
END_VAR

VAR
	_Member	: KOSTAL_AF2024_Core_System.I_Interface;
END_VAR

//preset
IF 		__ISVALIDREF(rFound_I)	THEN	rFound_I:= _Dummy;	
ELSE 	_setResultFail(Response, "no reference to rFound_I found");	RETURN;  
END_IF	

IF Number = 0 THEN _setResultFail(Response, "Number is out of range (1..n)"); RETURN; END_IF

IF _findMemberByIndex(Number - 1, _Member, Response) THEN
	Get_I:= _get_I(_Member, rFound_I, Response);
END_IF
END_METHOD

(*
	Get full access to content of Member with {Number}
*) 
METHOD Get_I_Owner : BOOL

VAR_INPUT
	Number		: UDINT;
	rFound_I	: REFERENCE TO I_T_Tool_Owner;
	Response	: KOSTAL_AF2024_Core_functionResponse.I_T_functionResponse_Owner;
END_VAR

VAR
	_Member	: KOSTAL_AF2024_Core_System.I_Interface;
END_VAR

//preset
IF 		__ISVALIDREF(rFound_I)	THEN	rFound_I:= _Dummy;	
ELSE 	_setResultFail(Response, "no reference to rFound_I found");	RETURN;  
END_IF	

IF Number = 0 THEN _setResultFail(Response, "Number is out of range (1..n)"); RETURN; END_IF

IF _findMemberByIndex(Number - 1, _Member, Response) THEN
	Get_I_Owner:= _get_I_Owner(_Member, rFound_I, Response);
END_IF
END_METHOD

(*
	Number of Member in list.
*)
PROPERTY NumberOfMember : UDINT
GET

NumberOfMember:= SUPER^._NumberOfMember;
END_GET
END_PROPERTY

END_FUNCTION_BLOCK

// TcpIp/DUT/Tool/T_Tool
{attribute 'enable_dynamic_creation'}
(*
	Example class for use within a list.
	Make sure that the atrribute shown above is present in your class in this form and location.
*)
FUNCTION_BLOCK T_Tool IMPLEMENTS I_T_Tool, I_T_Tool_CopyFrom, I_T_Tool_Owner

VAR
	_Number			:	UINT;
	_Pass				:	BOOL;
	_MatchingRate	: KOSTAL_AF2024_Core_Settings.T_MaxString_UTF8;
END_VAR

METHOD PUBLIC Clear

_Number	:= 0;
_Pass		:= FALSE;
END_METHOD

METHOD PUBLIC CopyFrom : BOOL
VAR_INPUT
	IN	: KOSTAL_AF2024_Core_System.I_Interface;
END_VAR


VAR
	_obj		: I_T_Tool_Owner;
	_obj2		: I_T_Tool;
END_VAR

Clear();

IF IN = 0 THEN RETURN;

ELSIF __QUERYINTERFACE(IN, _obj) AND_THEN _obj <> 0 THEN

	_Number			:= _obj.Number;
	_Pass				:= _obj.Pass;
	_MatchingRate	:= _obj.MatchingRate;

	CopyFrom:= TRUE;
	
ELSIF __QUERYINTERFACE(IN, _obj2) AND_THEN _obj2 <> 0 THEN

	_Number			:= _obj2.Number;
	_Pass				:= _obj2.Pass;
	_MatchingRate	:= _obj2.MatchingRate;

	CopyFrom:= TRUE;
	
END_IF
END_METHOD

METHOD PUBLIC CopyTo : bool
VAR_INPUT
	IN	: I_T_Tool_CopyFrom;
END_VAR

IF IN = 0 THEN RETURN;	END_IF

CopyTo:= IN.CopyFrom(THIS^);
END_METHOD

PROPERTY PUBLIC MatchingRate : KOSTAL_AF2024_Core_Settings.T_MaxString_UTF8
GET

MatchingRate:= _MatchingRate;
END_GET
SET

_MatchingRate:= MatchingRate;
END_SET
END_PROPERTY

PROPERTY PUBLIC Number : UINT
GET

Number:= _Number;
END_GET
SET

_Number:= Number;
END_SET
END_PROPERTY

PROPERTY PUBLIC Pass : BOOL
GET

Pass:= _Pass;
END_GET
SET

_Pass:= Pass;
END_SET
END_PROPERTY

END_FUNCTION_BLOCK

// TcpIp/DUT/Version/I_T_SensorVersion_TcpIp
INTERFACE I_T_SensorVersion_TcpIp EXTENDS KOSTAL_AF2024_Core_System.I_Interface

METHOD PUBLIC CopyTo : BOOL
VAR_INPUT
	IN	: I_T_SensorVersion_TcpIp_CopyFrom;
END_VAR
END_METHOD

PROPERTY PUBLIC HeadModel : KOSTAL_AF2024_Core_Settings.T_MaxString_UTF8
GET
END_GET
END_PROPERTY

PROPERTY PUBLIC Version : KOSTAL_AF2024_Core_Settings.T_MaxString_UTF8
GET
END_GET
END_PROPERTY

END_INTERFACE

// TcpIp/DUT/Version/I_T_SensorVersion_TcpIp_CopyFrom
INTERFACE I_T_SensorVersion_TcpIp_CopyFrom EXTENDS KOSTAL_AF2024_Core_System.I_Interface

METHOD PUBLIC CopyFrom : BOOL
VAR_INPUT
	IN	: I_T_SensorVersion_TcpIp;
END_VAR
END_METHOD

END_INTERFACE

// TcpIp/DUT/Version/I_T_SensorVersion_TcpIp_Owner
INTERFACE I_T_SensorVersion_TcpIp_Owner EXTENDS I_T_SensorVersion_TcpIp

METHOD PUBLIC Clear
VAR_INPUT
END_VAR
END_METHOD

METHOD PUBLIC CopyFrom : BOOL
VAR_INPUT
	IN	: I_T_SensorVersion_TcpIp;
END_VAR
END_METHOD

PROPERTY PUBLIC HeadModel : KOSTAL_AF2024_Core_Settings.T_MaxString_UTF8
SET
END_SET
END_PROPERTY

PROPERTY PUBLIC Version : KOSTAL_AF2024_Core_Settings.T_MaxString_UTF8
SET
END_SET
END_PROPERTY

END_INTERFACE

// TcpIp/DUT/Version/T_SensorVersion_TcpIp
FUNCTION_BLOCK PUBLIC T_SensorVersion_TcpIp IMPLEMENTS I_T_SensorVersion_TcpIp, I_T_SensorVersion_TcpIp_Owner, I_T_SensorVersion_TcpIp_CopyFrom
VAR
	_HeadModel	: KOSTAL_AF2024_Core_Settings.T_MaxString_UTF8;
	_Version		: KOSTAL_AF2024_Core_Settings.T_MaxString_UTF8;
END_VAR

METHOD PUBLIC Clear
VAR_INPUT
END_VAR

_HeadModel	:= '';
_Version		:= '';
END_METHOD

METHOD PUBLIC CopyFrom : BOOL
VAR_INPUT
	IN	: I_T_SensorVersion_TcpIp;
END_VAR

VAR
	_obj	: I_T_SensorVersion_TcpIp;
END_VAR

IF (IN = 0) OR_ELSE NOT __QUERYINTERFACE(IN, _obj) OR_ELSE (_obj = 0) THEN RETURN;	END_IF

_HeadModel	:= IN.HeadModel;
_Version		:= IN.Version;

CopyFrom:= TRUE;
END_METHOD

METHOD PUBLIC CopyTo : BOOL
VAR_INPUT
	IN	: I_T_SensorVersion_TcpIp_CopyFrom;
END_VAR

VAR
	_obj	: I_T_SensorVersion_TcpIp_CopyFrom;
END_VAR

IF (IN = 0) OR_ELSE NOT __QUERYINTERFACE(IN, _obj) OR_ELSE (_obj = 0) THEN RETURN;	END_IF

CopyTo:= IN.CopyFrom(THIS^);
END_METHOD

PROPERTY PUBLIC HeadModel : KOSTAL_AF2024_Core_Settings.T_MaxString_UTF8
GET

HeadModel:= _HeadModel;
END_GET
SET

_HeadModel:= HeadModel;
END_SET
END_PROPERTY

PROPERTY PUBLIC Version : KOSTAL_AF2024_Core_Settings.T_MaxString_UTF8
GET

Version:= _Version;
END_GET
SET

_Version:= Version;
END_SET
END_PROPERTY

END_FUNCTION_BLOCK

// TcpIp/FB_Camera_TcpIp_IV
FUNCTION_BLOCK PUBLIC FB_Camera_TcpIp_IV IMPLEMENTS I_Camera_TcpIp_IV
VAR CONSTANT
		_PortDefault	: UDINT:= 8500;
		_MaxPrg				: UDINT:= 127;
END_VAR

VAR
	_serverAmsNetId	: Tc2_System.T_AmsNetID:= '';
	_IP							: Tc2_System.T_IPv4Addr;
	_Port						: UDINT:= _PortDefault;

	_socket								: Tc2_TcpIp.FB_ClientServerConnection;
	_executedSocketState	:	Tc2_TcpIp.E_SocketConnectionState;
	
	_send						: Tc2_TcpIp.FB_SocketSend;
	_receive				: Tc2_TcpIp.FB_SocketReceive;

	_receivedPartly	: KOSTAL_AF2024_Core_Settings.T_MaxString_UTF8;

	_COMMAND_TCPIP	: _T_Command;
	
	_Command	: KOSTAL_AF2024_Core_Settings.T_MaxString_UTF8:= '||0:000>TRIGGER ON$0D$0A';	//default
	_ETX									: STRING(1):= '$0D';	//Carriage Return
	_intermediateLimiter	: STRING(1):= '$2C';	//comma

	_timeOut			: TIME	:= T#5S;	//default T#5S
	_timeOutTimer	: TON;	//TON

	_ProgramNumber		: UINT;
	_ProgramNumberGet	: UINT;
	
	_receivedString	: KOSTAL_AF2024_Core_Settings.T_MaxString_UTF8;
	_split					: KOSTAL_AF2024_Core_StringTools.FB_Split_UTF8;
	_responses			: KOSTAL_AF2024_Core_ListOf.FB_ListOfString_UTF8;
	
	_Step					: KOSTAL_AF2024_Core_Process.FB_processStep;
	_SubStep			: KOSTAL_AF2024_Core_Process.FB_processStep;
	_Init					: BOOL:= TRUE;
	_PrepareCycle	: BOOL;	//Set {_PrepareCycle} to suppress a finish state in this cycle.
	
	_state		:	KOSTAL_AF2024_Core_Process.T_plcState;


	_THIS_CALLED			: _E_THIS_TcpIp;
	_THIS_IN_PROCESS	: _E_THIS_TcpIp;

	//_LastResult	: BOOL;
	_Version		:	T_SensorVersion_TcpIp;
	_Result_RT	: T_Response_RT_TcpIp;

	_OpMode	: E_OpMode_TcpIp;

	_ErrorMessage	: KOSTAL_AF2024_Core_Settings.T_MaxString_UTF8;
END_VAR

VAR CONSTANT
	_ADDRESS_IDLE					: INT:= 0;
	_ADDRESS_SEND					: INT:= 1;

	_ADDRESS_TRIGGER_PRG	: INT:= 100;
END_VAR

METHOD FB_init : BOOL
VAR_INPUT
	bInitRetains : BOOL; // if TRUE, the retain variables are initialized (warm start / cold start)
	bInCopyCode : BOOL;  // if TRUE, the instance afterwards gets moved into the copy code (online change)
	AmsNetId		: Tc2_System.T_AmsNetID;	//AmsNetId from system which provides the TcpIp Server
	IP					: Tc2_System.T_IPv4Addr;	//Camera IP address
	Port				: UDINT;									//Camera port
END_VAR

IF AmsNetId <> ''	THEN	_serverAmsNetId:= AmsNetId;	END_IF
IF IP <> ''				THEN	_IP:= IP;										END_IF
IF Port	<> 0			THEN	_Port:= Port;								END_IF
END_METHOD

METHOD PROTECTED _getCommand : KOSTAL_AF2024_Core_Settings.T_MaxString_UTF8

VAR_INPUT
	ID				: _E_Command_TcpIp;
	Parameter : UINT;
END_VAR
VAR
	_c	: KOSTAL_AF2024_Core_StringTools.FB_Concat_UTF8;
	_s	: KOSTAL_AF2024_Core_Settings.T_MaxString_UTF8;
END_VAR

CASE ID OF
	
	_E_Command_TcpIp.Trigger						: _getCommand:= _mergePlCommand(_COMMAND_TCPIP.TriggerAndState);
	_E_Command_TcpIp.GetProgram				:	_getCommand:= _mergePlCommand(_COMMAND_TCPIP.GetProgram); 
	_E_Command_TcpIp.ReadVersion				:	_getCommand:= _mergePlCommand(_COMMAND_TCPIP.ReadVersion);
	_E_Command_TcpIp.ReadOperationMode	:	_getCommand:= _mergePlCommand(_COMMAND_TCPIP.ReadOperationMode);

	_E_Command_TcpIp.SetProgram	:	_c.clear(); _c.addContent(_COMMAND_TCPIP.SetProgram);			_c.addContent(',');
																_c.addContent(KOSTAL_AF2024_Core_StringTools.F_FormatMask_UTF8(TO_STRING(Parameter), '000', KOSTAL_AF2024_Core_StringTools.E_ALIGNMENT.RIGHT));
																_c.addContent(_ETX); _getCommand:= _c.getResult(); _c.clear();


END_CASE
END_METHOD

//mergeParameterlessCommand - return a commandstring without additional input parameters
METHOD PROTECTED _mergePlCommand : KOSTAL_AF2024_Core_Settings.T_MaxString_UTF8
VAR_INPUT
	Command		: KOSTAL_AF2024_Core_Settings.T_MaxString_UTF8;
END_VAR

VAR
	_c	: KOSTAL_AF2024_Core_StringTools.FB_Concat_UTF8;
END_VAR

_c.Clear(); 
_c.addContent(Command);	
//_c.addContent(',');	
_c.addContent(_ETX); 
_mergePlCommand:= _c.getResult();	
_c.Clear();
END_METHOD

METHOD PROTECTED _Parse_Error : BOOL
VAR_INPUT
	IN	: _E_THIS_TcpIp;
END_VAR

VAR
	_c: KOSTAL_AF2024_Core_StringTools.FB_Concat_UTF8;
END_VAR

IF _responses.line_GET(1) = _COMMAND_TCPIP.Error THEN

	_Parse_Error:= TRUE;
	
	IF _Step.toggle THEN	_Parse_ErrorMessage(IN);	END_IF
	
	_state.clear();
	_state.finish:= TRUE;
	_state.fail:= TRUE;
	_state.description:= TO_WSTRING(_ErrorMessage);

END_IF
END_METHOD

METHOD PROTECTED _Parse_ErrorMessage
VAR_INPUT
	IN	: _E_THIS_TcpIp;
END_VAR

VAR
	_c: KOSTAL_AF2024_Core_StringTools.FB_Concat_UTF8;
	_fErr: UINT;
END_VAR

_ErrorMessage:= 'ERROR;Code:';

_c.Clear();
_c.addContent(_responses.line_GET(3));
_c.addContent(';');


CASE IN OF
	
	_E_THIS_TcpIp.GetProgram		:	_c.addContent('Get Programm[');	
	_E_THIS_TcpIp.SetProgram		:	_c.addContent('Set Programm[');	
	_E_THIS_TcpIp.Trigger			:	_c.addContent('Trigger[');	
	_E_THIS_TcpIp.TriggerPrgNo	:	_c.addContent('TriggerPrg[');	
	_E_THIS_TcpIp.ReadVersion	:	_c.addContent('Read Version[');	

ELSE													_c.addContent('Unknown Command[');
END_CASE

_c.addContent(_responses.line_GET(2));
_c.addContent('];');

_fErr	:= TO_UINT(_responses.line_GET(3));

CASE _fErr OF
	0	: _c.addContent('no Error');

	1..32 :	_c.addContent('Program number ');
					_c.addContent(_responses.line_GET(2));
					_c.addContent(' Error Damage');
	
	52 :	_c.addContent('Program switching error(commissioning;external input)');
	53 :	_c.addContent('Program switching error (commissioning; panel/PC/network)');
	75 :	_c.addContent('Non-volatile memory error (EEPROM)');
	76 :	_c.addContent('Non-volatile memory error (FLASHROM)');
	79 :	_c.addContent('Program switching error (runtime)');
	81..123,125..128 :	_c.addContent('System error. It is possible that an error has occurred inside the sensor.');
	124 :	_c.addContent('System error. No sensor head is connected to the evaluation unit.');

	ELSE _c.addContent('no definition found for this error code');
END_CASE

_ErrorMessage:= _c.getResult();

_c.clear();
END_METHOD

METHOD PROTECTED _Parse_GetProgram

IF _step.toggle THEN

	
	_state.clear();
	
	IF _responses.line_GET(1) <> _COMMAND_TCPIP.GetProgram THEN

		_state.finish:= TRUE;
		_state.fail:= TRUE;
		_state.description:= "The command was NOT returned correctly.";

	ELSE

		_ProgramNumberGet	:= TO_UINT(_responses.line_GET(2));
		
		_Step.INC();

	END_IF		

END_IF
END_METHOD

METHOD PROTECTED _Parse_OpMode

IF _step.toggle THEN

	
	_state.clear();
	
	IF _responses.line_GET(1) <> _COMMAND_TCPIP.ReadOperationMode THEN

		_state.finish:= TRUE;
		_state.fail:= TRUE;
		_state.description:= "The command was NOT returned correctly.";

	ELSE

		IF 		TO_UINT(_responses.line_GET(2)) = 0 THEN	_OpMode:= E_OpMode_TcpIp.Setup;
		ELSIF TO_UINT(_responses.line_GET(2)) = 1 THEN	_OpMode:= E_OpMode_TcpIp.Run;
		ELSE 																						_OpMode:= E_OpMode_TcpIp.Unknown;
		END_IF		

		_Step.INC();

	END_IF		

END_IF
END_METHOD

METHOD PROTECTED _Parse_SetProgram

IF _step.toggle THEN

	
	_state.clear();
	
	IF _responses.line_GET(1) <> _COMMAND_TCPIP.SetProgram THEN

		_state.finish:= TRUE;
		_state.fail:= TRUE;
		_state.description:= "The command was NOT returned correctly.";

	ELSE

		_Step.INC();

	END_IF		

END_IF
END_METHOD

METHOD PROTECTED _Parse_Trigger


VAR
	_udi	: UDINT;
	_tool	: T_Tool;
END_VAR

IF _step.toggle THEN

	
	_state.clear();
	
	IF _responses.line_GET(1) <> _COMMAND_TCPIP.StateResult THEN

		_state.finish:= TRUE;
		_state.fail:= TRUE;
		_state.description:= "The command was NOT returned correctly.";

	ELSIF (_responses.NumberOfLines - 3) MOD 3 <> 0 THEN 

		_state.finish:= TRUE;
		_state.fail:= TRUE;
		_state.description:= "Tools are not returned correctly";

	ELSE

		_Result_RT.ResultCount	:= TO_UDINT(_responses.line_GET(2));
		_Result_RT.OverallPass	:= _responses.line_GET(3) = _COMMAND_TCPIP.OK;
		
		FOR _udi:= 4 TO _responses.NumberOfLines BY 3 DO
			_tool.Clear();
			_tool.Number			:= TO_UINT(_responses.line_GET(_udi));
			_tool.Pass				:= _responses.line_GET(_udi + 1) = _COMMAND_TCPIP.OK;
			_tool.MatchingRate	:= _responses.line_GET(_udi + 2);
			_Result_RT.Tools_Owner.Add_DUT(_tool, 0);
		END_FOR

		_tool.Clear();
		
		_Step.INC();

	END_IF		

END_IF
END_METHOD

METHOD PROTECTED _Parse_Version

IF _step.toggle THEN

	
	_state.clear();
	
	IF _responses.line_GET(1) <> _COMMAND_TCPIP.ReadVersion THEN

		_state.finish:= TRUE;
		_state.fail:= TRUE;
		_state.description:= "The command was NOT returned correctly.";

	ELSE

		_Version.HeadModel	:= _responses.line_GET(2);
		_Version.Version		:= _responses.line_GET(3);
		
		_Step.INC();

	END_IF		

END_IF
END_METHOD

METHOD PROTECTED _a0_stepFail
VAR_INPUT
END_VAR

	_state.clear();
	_state.description:= Tc2_Standard.WCONCAT("Step does not exist: ", INT_TO_WSTRING(_step.actual));
	_state.fail		:= TRUE;
	_state.finish	:= TRUE;
END_METHOD

METHOD PUBLIC _a0_stepInit
VAR_INPUT
END_VAR

//Overwrite base method

IF _Init THEN

	_step.init();
	_Init:= FALSE;	

	_socket.bEnable		:= FALSE;
	_send.bExecute		:= FALSE;
	_receive.bExecute	:= FALSE;

	_timeOutTimer.IN:= FALSE;

ELSIF _THIS_CALLED <> _THIS_IN_PROCESS AND _step.actual > 0 THEN 

	_step.init();

	_socket.bEnable		:= FALSE;
	_send.bExecute		:= FALSE;
	_receive.bExecute	:= FALSE;

	_timeOutTimer.IN:= FALSE;

END_IF
END_METHOD

METHOD PROTECTED _a1_Finish
VAR_INPUT
END_VAR

IF _step.toggle THEN

	_timeOutTimer.IN:= FALSE;

	_socket.bEnable		:= FALSE;
	_send.bExecute		:= FALSE;
	_receive.bExecute	:= FALSE;

END_IF

IF _PrepareCycle THEN	_Step.set(_ADDRESS_IDLE);
ELSE
	_state.clear();
	_state.finish	:= TRUE;
	_state.pass		:= TRUE;
END_IF
END_METHOD

METHOD PROTECTED _a1_Idle
VAR_INPUT
END_VAR

_state.clear();

_THIS_IN_PROCESS:= _E_THIS_TcpIp.Idle;


IF _step.toggle THEN

	_socket(bEnable		:= FALSE);
	_send(bExecute		:= FALSE);
	_receive(bExecute	:= FALSE);

	_timeOutTimer(IN:= FALSE);

	_state.busy:= TRUE;

	
ELSIF 	_socket.bBusy THEN

	_state.busy:= TRUE;
	_state.description:= "socket is busy, please wait...";
	
ELSIF _send.bBusy THEN

	_state.busy:= TRUE;
	_state.description:= "send is busy, please wait...";

	
ELSIF _receive.bBusy THEN

	_state.busy:= TRUE;
	_state.description:= "receive is busy, please wait...";

ELSIF _THIS_CALLED = _E_THIS_TcpIp.Idle THEN

	_state.ready:= TRUE;

	
ELSIF _THIS_CALLED = _E_THIS_TcpIp.Trigger THEN

	
	_THIS_IN_PROCESS:= _THIS_CALLED;

	_state.busy:= TRUE;

	_receivedString:= '';
	_receivedPartly:= '';
	
	_split.clear();
	_responses.clear();
	
	_timeOutTimer.IN:= TRUE;
	
	_state.clear();
	_state.busy:= TRUE;

	_Result_RT.Clear();
	
	_Command	:= _getCommand(_E_Command_TcpIp.Trigger, 0);

	_step.set(_ADDRESS_SEND);
	
	
ELSIF _THIS_CALLED = _E_THIS_TcpIp.TriggerPrgNo THEN

	
	_THIS_IN_PROCESS:= _THIS_CALLED;

	_state.busy:= TRUE;

	_receivedString:= '';
	_receivedPartly:= '';
	
	_split.clear();
	_responses.clear();
	_Result_RT.Clear();
	
	_timeOutTimer.IN:= TRUE;
	
	_state.clear();
	_state.busy:= TRUE;

	_step.set(_ADDRESS_TRIGGER_PRG);
	
	

ELSIF _THIS_CALLED = _E_THIS_TcpIp.SetProgram THEN


	_THIS_IN_PROCESS:= _THIS_CALLED;

	IF _Programnumber > _MaxPrg THEN
		
		_state.description:= "Number of program is out of range (0..127)";
		_state.fail:= TRUE;
		_state.finish:= TRUE;

	ELSE

		_state.busy:= TRUE;
	
		_timeOutTimer.IN:= TRUE;
		
		_state.clear();
		_state.busy:= TRUE;

		_Command	:= _getCommand(_E_Command_TcpIp.SetProgram, _ProgramNumber);

		_step.set(_ADDRESS_SEND);
		
	END_IF
	
	
ELSIF _THIS_CALLED = _E_THIS_TcpIp.GetProgram THEN

	_THIS_IN_PROCESS:= _THIS_CALLED;

	IF _ProgramNumber > _MaxPrg THEN
		
		_state.description:= "Number of program is out of range (0..127)";
		_state.fail:= TRUE;
		_state.finish:= TRUE;

	ELSE

		_state.busy:= TRUE;
	
		_timeOutTimer.IN:= TRUE;
		
		_state.clear();
		_state.busy:= TRUE;

		_Command	:= _getCommand(_E_Command_TcpIp.GetProgram, 0);

		_step.set(_ADDRESS_SEND);
		
	END_IF

ELSIF _THIS_CALLED = _E_THIS_TcpIp.ReadVersion THEN

	_THIS_IN_PROCESS:= _THIS_CALLED;

	_state.busy:= TRUE;

	_timeOutTimer.IN:= TRUE;
	
	_state.clear();
	_state.busy:= TRUE;

	_Version.Clear();
	
	_Command	:= _getCommand(_E_Command_TcpIp.ReadVersion, 0);

	_step.set(_ADDRESS_SEND);
		
ELSIF _THIS_CALLED = _E_THIS_TcpIp.ReadOperationMode THEN

	_THIS_IN_PROCESS:= _THIS_CALLED;

	_state.busy:= TRUE;

	_timeOutTimer.IN:= TRUE;
	
	_state.clear();
	_state.busy:= TRUE;

	_OpMode:= E_OpMode_TcpIp.Unknown;
	
	_Command	:= _getCommand(_E_Command_TcpIp.ReadOperationMode, 0);

	_step.set(_ADDRESS_SEND);
		

ELSE

	_state.clear();
	_state.ready:= TRUE;
		
END_IF
END_METHOD

METHOD PROTECTED _a2_Connect
VAR
	_c	: KOSTAL_AF2024_Core_StringTools.FB_Concat;
END_VAR

IF _step.toggle THEN
	_state.clear();
	_state.busy:= TRUE;
	_subStep.init();
END_IF


IF _timeOutTimer.Q THEN

	_timeOutOccured();

ELSE

	_subStep.Header();
	
	CASE _subStep.actual OF
		0:	_socket.bEnable:= FALSE;	_subStep.INC();
		1:	_socket.bEnable:= TRUE;		_subStep.INC();

		2:	IF _socket.bBusy THEN
					_state.busy	:= TRUE;
					_state.description:= "Scanner is busy(connect); wait ...";
				ELSE
					_subStep.INC();
				END_IF

		3:	IF _socket.bError THEN
					_state.clear();
					_state.description:= Tc2_Standard.WCONCAT("Error during socket open. Errorcode>", UDINT_TO_WSTRING(_socket.nErrId));
					_state.fail	:= TRUE;
					_state.finish:= TRUE;	
					_timeOutTimer.IN:= FALSE;
				ELSIF _socket.hSocket.handle = 0 THEN
					_state.clear();
					_state.description:= "no Handle from socket";
					_state.fail	:= TRUE;
					_state.finish:= TRUE;
					_timeOutTimer.IN:= FALSE;
				ELSE
					_step.INC();
				END_IF
		
	ELSE
	
		_timeOutTimer.IN:= FALSE;
		_state.clear();
		_state.fail	:= TRUE;
		_state.finish:= TRUE;
		_c.clear();
		_c.addContent("connect Step ");
		_c.addContent(INT_TO_WSTRING(_subStep.actual));
		_c.addContent(" does not exist");
		_state.description:= _c.getResult();
		_c.clear();
	
	END_CASE

END_IF
END_METHOD

METHOD PROTECTED _a2_Parse
VAR_INPUT
	IN	: _E_THIS_TcpIp;
END_VAR

IF _Parse_Error(IN) THEN RETURN;	END_IF

CASE IN OF
	
	_E_THIS_TcpIp.Idle :	_step.INC();	//no parsing available

	_E_THIS_TcpIp.ReadVersion				:	_Parse_Version();
	_E_THIS_TcpIp.Trigger 						:	_Parse_Trigger();
	_E_THIS_TcpIp.TriggerPrgNo				:	_Parse_Trigger();
	_E_THIS_TcpIp.GetProgram					:	_Parse_GetProgram();
	_E_THIS_TcpIp.SetProgram					:	_Parse_SetProgram();
	_E_THIS_TcpIp.ReadOperationMode	:	_Parse_OpMode();
	
END_CASE
END_METHOD

METHOD PROTECTED _a2_Receive
VAR
	_c	: KOSTAL_AF2024_Core_StringTools.FB_Concat;
END_VAR

IF _step.toggle THEN

	_state.clear();
	_state.busy:= TRUE;

	_subStep.init();

	_receivedString:= '';
	_receivedPartly:= '';

	_split.clear();
	_responses.clear();

END_IF



IF _timeOutTimer.Q THEN

	_timeOutOccured();

ELSE
	
	_subStep.Header();

	CASE _subStep.actual OF

		0:	_receive.bExecute:= FALSE;	_receivedPartly:= '';	_subStep.INC();
		1:	_receive.bExecute:= TRUE;		_subStep.INC();

		2:	IF _receive.bBusy THEN
					_state.busy	:= TRUE;
					_state.description:= "Scanner is busy(receive); wait ...";
				ELSE
					_subStep.INC();
				END_IF

		3:	IF _receive.bError THEN
					_state.clear();
					_state.description:= Tc2_Standard.WCONCAT("Error during receive. Errorcode>", UDINT_TO_WSTRING(_receive.nErrId));
					_state.fail	:= TRUE;
					_state.finish:= TRUE;	
					_timeOutTimer.IN:= FALSE;
				ELSE
					_subStep.INC();
				END_IF
		
		4:	IF	_receive.nRecBytes <> 0 THEN 

					_receivedString:= Tc2_Standard.CONCAT(STR1:= _receivedString, STR2:=  Tc2_Standard.LEFT(STR:= _receivedPartly, SIZE:= UDINT_TO_INT(_receive.nRecBytes)));
					_receivedPartly:= '';

					IF NOT _splitString() THEN	_subStep.SET(0);
					ELSE
						_state.clear();
						_state.busy:= TRUE;
						_state.pass:= TRUE;
						_timeOutTimer.IN:= FALSE;
						_step.INC();
					END_IF
					
				ELSE	_subStep.SET(0);

				END_IF
								
	ELSE
	
		_timeOutTimer.IN:= FALSE;
		_state.clear();
		_state.fail	:= TRUE;
		_state.finish:= TRUE;
		_c.clear();
		_c.addContent("send Step ");
		_c.addContent(INT_TO_WSTRING(_subStep.actual));
		_c.addContent(" does not exist");
		_state.description:= _c.getResult();
		_c.clear();
	
	END_CASE

END_IF
END_METHOD

METHOD PROTECTED _a2_Send
VAR
	_c	: KOSTAL_AF2024_Core_StringTools.FB_Concat;
END_VAR

IF _step.toggle THEN
	_state.clear();
	_state.busy:= TRUE;
	_subStep.init();
END_IF


IF _timeOutTimer.Q THEN

	_timeOutOccured();

ELSE
	
	_subStep.Header();

	CASE _subStep.actual OF
		0:	_send.bExecute:= FALSE;	_subStep.INC();
		1:	_send.bExecute:= TRUE;		_subStep.INC();

		2:	IF _send.bBusy THEN
					_state.busy	:= TRUE;
					_state.description:= "Scanner is busy(send); wait ...";
				ELSE
					_subStep.INC();
				END_IF

		3:	IF _send.bError THEN
					_state.clear();
					_state.description:= Tc2_Standard.WCONCAT("Error during send. Errorcode>", UDINT_TO_WSTRING(_send.nErrId));
					_state.fail	:= TRUE;
					_state.finish:= TRUE;	
					_timeOutTimer.IN:= FALSE;
				ELSE
					_step.INC();
				END_IF
		
	ELSE
	
		_state.clear();
		_state.fail	:= TRUE;
		_state.finish:= TRUE;
		_c.clear();
		_c.addContent("send Step ");
		_c.addContent(INT_TO_WSTRING(_subStep.actual));
		_c.addContent(" does not exist");
		_state.description:= _c.getResult();
		_c.clear();
	
	END_CASE

END_IF
END_METHOD


METHOD PROTECTED _a3_PrgIsEqual
VAR_INPUT
END_VAR

//if get program same as set requested program call trgger 

IF _Step.toggle THEN	;	END_IF

IF _ProgramNumber = _ProgramNumberGet THEN	

	_Command	:= _getCommand(_E_Command_TcpIp.Trigger, 0);	_Step.INC();
	_Step.set(_ADDRESS_SEND);

ELSE	_Step.INC();
	
END_IF
END_METHOD

METHOD PROTECTED _devices
VAR_INPUT
END_VAR


_timeOutTimer(IN:= , PT:= _timeOut, Q=> , ET=> );

_socket
	(
		sSrvNetID	:= _serverAmsNetId, 
		nMode			:= Tc2_TcpIp.CONNECT_MODE_ENABLEDBG, 

		sRemoteHost	:= _IP, 
		nRemotePort	:= _Port, 

		bEnable			:= , 
		tReconnect	:= _timeOut, 

		bBusy		=> , 
		bError	=> , 
		nErrId	=> , 
		hSocket	=> , 
		eState	=> 
	);
	
IF _socket.bEnable THEN	_executedSocketState:= _socket.eState;	END_IF
	
_send
	(
		sSrvNetId	:= _serverAmsNetId, 
		hSocket		:= _socket.hSocket, 
		cbLen			:= SIZEOF(_Command), 
		pSrc			:= ADR(_Command), 
		bExecute	:= , 
		tTimeout	:= _timeOut, 

		bBusy			=> , 
		bError		=> , 
		nErrId		=> 
	);
	
	
	_receive
	(
		sSrvNetId	:= _serverAmsNetId, 
		hSocket		:= _socket.hSocket, 

		cbLen:= SIZEOF(_receivedPartly) - 1, 
		pDest:= ADR(_receivedPartly), 

		bExecute:= , 
		tTimeout:= _timeOut, 

		bBusy			=> , 
		bError		=> , 
		nErrId		=> , 
		nRecBytes	=> 
	);
END_METHOD

(*
| split received string depends of STX ETX
*)
METHOD PROTECTED _splitString  : BOOL

VAR
	_udi: UDINT;
	_element: KOSTAL_AF2024_Core_Settings.T_MaxString_UTF8;
	_stxPos: INT;
	_code			: KOSTAL_AF2024_Core_Settings.T_MaxString_UTF8;
END_VAR
_responses.clear();

_stxPos:= Tc2_Standard.FIND(_receivedString, _ETX);

IF 		_stxPos = 0 THEN	;	// no splitting possible
ELSIF _stxPos = 1 THEN	_splitString:= TRUE;	// response is empty
ELSE	

	_code:= Tc2_System.LEFT(_receivedString, _stxPos - 1);
	
	_split.clear();
	_split.Delimiter:= _intermediateLimiter;
	_split.split(_code);

	FOR _udi:= 1 TO _split.Results.NumberOfLines DO
		_responses.addLine(newLine:= _split.Results.line_GET(_udi));
	END_FOR

	_splitString:= TRUE;	

END_IF
END_METHOD

METHOD PROTECTED _timeOutOccured
VAR_INPUT
END_VAR


_socket.bEnable		:= FALSE;
_send.bExecute		:= FALSE;
_receive.bExecute	:= FALSE;

_state.busy:= FALSE;
_state.description:= "Timeout";
_state.fail:= TRUE;
_state.finish:= TRUE;
END_METHOD

(*
Decription
==========
*)
METHOD PROTECTED _FBmain


_a0_stepInit();

_step.Header();

CASE _step.actual OF

	_ADDRESS_IDLE:	_a1_Idle();

	_ADDRESS_SEND:	_a2_Connect();
	2:	_a2_Send();
	3:	_a2_Receive();
	4:	_a2_Parse(_THIS_IN_PROCESS);
	5:	_a1_Finish();

	_ADDRESS_TRIGGER_PRG:		
				_Command	:= _getCommand(_E_Command_TcpIp.GetProgram, 0);	_Step.INC();
	101:	_a2_Connect();
	102:	_a2_Send();
	103:	_a2_Receive();
	104:	_a2_Parse(_E_THIS_TcpIp.GetProgram);

	105:	_a3_PrgIsEqual();

	106:	_Command	:= _getCommand(_E_Command_TcpIp.SetProgram, _ProgramNumber);	_Step.INC();
	107:	_a2_Connect();
	108:	_a2_Send();
	109:	_a2_Receive();
	110:	_a2_Parse(_E_THIS_TcpIp.SetProgram);
	111:	_Command	:= _getCommand(_E_Command_TcpIp.Trigger, 0);		_Step.set(_ADDRESS_SEND);
	
	
(*
	_ADDRESS_SET_MAX_INDEX:	_IndexCounter:= 1;	 _step.INC();
	101:	_a2_Connect();
	102:	_a4_LoopHeader_MaxIndex(); 
	103:	_a2_Send();
	104:	_a4_LoopBottom();

	_ADDRESS_ENABLE_SETUP:	_step.INC();
	101:	_a2_Connect();
	102:	_a3_SelectSetup();
	103:	_a2_Send();
	104:	_a3_EnableSetup();
	105:	_a2_Send();
	106:	_a1_Finish();

	_ADDRESS_DISABLE_SETUP:	_step.INC();
	201:	_a2_Connect();
	202:	_a3_SelectSetup();
	203:	_a2_Send();
	204:	_a3_DisableSetup();
	205:	_a2_Send();
	206:	_a1_Finish();
*)

ELSE	_a0_stepFail();	

END_CASE
	
	

_devices();
END_METHOD

METHOD PUBLIC Clear

_responses.clear();
_receivedString:= '';
END_METHOD

METHOD PUBLIC Ex_GetProgramNumber : BOOL

VAR_INPUT
	ProgramNumber	: REFERENCE TO UINT;
END_VAR
IF _THIS_CALLED = _E_THIS_TcpIp.Idle THEN

	_THIS_CALLED:= _E_THIS_TcpIp.GetProgram;

	_FBmain();

	Ex_GetProgramNumber:= _THIS_CALLED = _THIS_IN_PROCESS;
	
	IF NOT __ISVALIDREF(ProgramNumber) THEN	;	//no valid reference
	ELSIF Ex_GetProgramNumber AND_THEN _state.finish AND_THEN _state.pass THEN ProgramNumber:= _ProgramNumberGet;	
	ELSE ProgramNumber:= 16#FFFF;	//no valid program number to response
	END_IF
	
ELSE
	
	Ex_GetProgramNumber:= FALSE;
 
END_IF
END_METHOD

METHOD PUBLIC Ex_ReadOperationMode : BOOL

VAR_INPUT
	OpMode	: REFERENCE TO E_OpMode_TcpIp;
END_VAR

IF _THIS_CALLED = _E_THIS_TcpIp.Idle THEN

	_THIS_CALLED:= _E_THIS_TcpIp.ReadOperationMode;

	_FBmain();

	Ex_ReadOperationMode:= _THIS_CALLED = _THIS_IN_PROCESS;

	IF NOT Ex_ReadOperationMode THEN	;
	ELSIF NOT __ISVALIDREF(OpMode) THEN 	;	//no valid reference
	ELSE OpMode:= _OpMode;
	END_IF
	
ELSE

	Ex_ReadOperationMode:= FALSE;
	
END_IF
END_METHOD

METHOD PUBLIC Ex_ReadVersion : BOOL

VAR_INPUT
	Version	: I_T_SensorVersion_TcpIp_Owner;
END_VAR

VAR
	_obj	: I_T_SensorVersion_TcpIp_Owner;
END_VAR

IF _THIS_CALLED = _E_THIS_TcpIp.Idle THEN

	_THIS_CALLED:= _E_THIS_TcpIp.ReadVersion;

	_FBmain();

	Ex_ReadVersion:= _THIS_CALLED = _THIS_IN_PROCESS;

	IF NOT Ex_ReadVersion THEN	;
	ELSIF (Version = 0) OR_ELSE NOT __QUERYINTERFACE(Version, _obj) OR_ELSE (_obj = 0) THEN 	;	//no valid reference
	ELSE Version.CopyFrom(_Version);
	END_IF
	
ELSE

	Ex_ReadVersion:= FALSE;
	
END_IF
END_METHOD

METHOD PUBLIC Ex_SetProgramNumber : BOOL

VAR_INPUT
	ProgramNumber	: UINT;
END_VAR
IF _THIS_CALLED = _E_THIS_TcpIp.Idle THEN

	_THIS_CALLED:= _E_THIS_TcpIp.SetProgram;

	_Programnumber:= ProgramNumber;

	_FBmain();

	Ex_SetProgramNumber:= _THIS_CALLED = _THIS_IN_PROCESS;
	
ELSE
	
	Ex_SetProgramNumber:= FALSE;
 
END_IF
END_METHOD

METHOD PUBLIC Ex_Trigger : BOOL

IF _THIS_CALLED = _E_THIS_TcpIp.Idle THEN

	_THIS_CALLED:= _E_THIS_TcpIp.Trigger;

	_FBmain();

	Ex_Trigger:= _THIS_CALLED = _THIS_IN_PROCESS;

ELSE

	Ex_Trigger:= FALSE;
	
END_IF
END_METHOD

METHOD PUBLIC Ex_Trigger_ProgramNumber : BOOL
VAR_INPUT
	ProgramNumber	: UINT;
END_VAR
IF _THIS_CALLED = _E_THIS_TcpIp.Idle THEN

	_THIS_CALLED:= _E_THIS_TcpIp.TriggerPrgNo;
	
	_ProgramNumber:= ProgramNumber;
	
	_FBmain();

	Ex_Trigger_ProgramNumber:= _THIS_CALLED = _THIS_IN_PROCESS;

ELSE

	Ex_Trigger_ProgramNumber:= FALSE;
	
END_IF
END_METHOD

METHOD PUBLIC GetElement : KOSTAL_AF2024_Core_Settings.T_MaxString_UTF8
VAR_INPUT
	number	: UINT;
END_VAR

GetElement:= _responses.line_GET(number);
END_METHOD

METHOD PUBLIC NativeStringGet : KOSTAL_AF2024_Core_Settings.T_MaxString_UTF8
VAR_INPUT
END_VAR

NativeStringGet:= _receivedString;
END_METHOD

(*
Description
===========
| IP address of the barcode reader
*)
PROPERTY PUBLIC IP : STRING
GET


IP:= _IP;
END_GET
SET

_IP:= IP;
END_SET
END_PROPERTY

(*
Description
===========
| TCP/IP port of the barcode reader
*)
PROPERTY PUBLIC Port : UDINT
GET


Port:= _Port;
END_GET
SET

IF Port = UDINT#0 THEN	_Port:= _PortDefault;
ELSE										_Port:= Port;
END_IF
END_SET
END_PROPERTY

PROPERTY PUBLIC Content : KOSTAL_AF2024_Core_ListOf.I_ListOfString_UTF8
GET

Content:= _responses;
END_GET
END_PROPERTY

(*
Description
===========
| State of the TCP/IP connection
*)
PROPERTY PUBLIC ExecutedSocketState : E_SocketConnectionState
GET

ExecutedSocketState:= _executedSocketState;
END_GET
END_PROPERTY

PROPERTY PUBLIC NumberOfEntries : UDINT
GET

NumberOfEntries:= _responses.NumberOfLines;
END_GET
END_PROPERTY

PROPERTY PUBLIC OperationMode : E_OpMode_TcpIp
GET

OperationMode:= _OpMode;
END_GET
END_PROPERTY

PROPERTY PUBLIC Result : I_T_Response_RT_TcpIp
GET

Result:= _Result_RT;
END_GET
END_PROPERTY

PROPERTY PUBLIC ResultPass : BOOL
GET

ResultPass:= _Result_RT.OverallPass;	//_LastResult;
END_GET
END_PROPERTY

(*
Description
===========
| AmsNetId of the system running the Beckhoff TCP/IP server
| default: ''=local system
*)
PROPERTY PUBLIC serverAmsNetId : STRING
GET

serverAmsNetId:= _serverAmsNetId;
END_GET
SET

_serverAmsNetId:= serverAmsNetId;
END_SET
END_PROPERTY

PROPERTY PUBLIC State : KOSTAL_AF2024_Core_Process.I_T_plcState
GET

State:= _state;
END_GET
END_PROPERTY

PROPERTY PUBLIC Version : I_T_SensorVersion_TcpIp
GET

Version:= _Version;
END_GET
END_PROPERTY

(*
Decription
==========
| To be called cyclicly, e.g. in DeviceDefine
*)
METHOD PUBLIC FBmain
VAR_INPUT
END_VAR

IF _THIS_CALLED = _E_THIS_TcpIp.Idle THEN
	_FBmain();
END_IF

_THIS_CALLED:= _E_THIS_TcpIp.Idle;
END_METHOD

END_FUNCTION_BLOCK

// TcpIp/I_Camera_TcpIp_IV
INTERFACE I_Camera_TcpIp_IV EXTENDS KOSTAL_AF2024_Drivers_Camera_I_Camera.I_Camera

METHOD PUBLIC GetElement : KOSTAL_AF2024_Core_Settings.T_MaxString_UTF8
VAR_INPUT
	number	: UINT;
END_VAR
END_METHOD

METHOD PUBLIC NativeStringGet : KOSTAL_AF2024_Core_Settings.T_MaxString_UTF8
VAR_INPUT
END_VAR
END_METHOD

PROPERTY PUBLIC Content : KOSTAL_AF2024_Core_ListOf.I_ListOfString_UTF8
GET
END_GET
END_PROPERTY

(*
Description
===========
| State of the TCP/IP connection
*)
PROPERTY PUBLIC ExecutedSocketState : E_SocketConnectionState
GET
END_GET
END_PROPERTY

(*
Description
===========
| IP address of the barcode reader
*)
PROPERTY PUBLIC IP : STRING
GET
END_GET
END_PROPERTY

PROPERTY PUBLIC NumberOfEntries : UDINT
GET
END_GET
END_PROPERTY

PROPERTY PUBLIC OperationMode : E_OpMode_TcpIp
GET
END_GET
END_PROPERTY

(*
Description
===========
| TCP/IP port of the barcode reader
*)
PROPERTY PUBLIC Port : UDINT
GET
END_GET
END_PROPERTY

PROPERTY PUBLIC Result : I_T_Response_RT_TcpIp
GET
END_GET
END_PROPERTY

(*
Description
===========
| AmsNetId of the system running the Beckhoff TCP/IP server
| default: ''=local system
*)
PROPERTY PUBLIC serverAmsNetId : STRING
GET
END_GET
END_PROPERTY

END_INTERFACE
